Staubli VAL3: initButton.pgx

public program initButton(utButton& x_utButton[], string x_sPage, string x_sId, string x_sText)
begin
  x_utButton.Common.sPage=x_sPage
  x_utButton.Common.sID=x_sId
  x_utButton.Common.sText=x_sText
  //
  //userPageBind(x_sPage,x_utButton.Common.sID,"style.backgroundColor",x_utButton.Appearance.sBackgroundColour,1,"r")
  userPageBind(x_utButton.Common.sPage,x_utButton.Common.sID,"innerHTML",x_utButton.Common.sText,1,"r")
  userPageBind(x_utButton.Common.sPage,x_utButton.Common.sID,"style.visibility",x_utButton.Appearance.bVisibility,1,"r")
  userPageBindClick(x_utButton.Common.sPage,x_utButton.Common.sID,x_utButton.Events.bClick,true)
  //
  x_utButton.Appearance.bVisibility=(x_sText!="")
  x_utButton.Events.bClick=false
end
